// TIA Portal V21 export
// export: Created 2026-11-21T23:19:43.1672142Z, ExportSetting WithDefaults, DisplayName Totally Integrated Automation Portal, DisplayVersion V21 Update 3, DisplayName STEP 7 Professional, DisplayVersion V21 Update 3, DisplayName STEP 7 Safety, DisplayVersion V21, DisplayName Tech WebApplication, DisplayVersion V21, DisplayName WinCC Basic/Comfort/Advanced, DisplayVersion V21 Update 3, DisplayName WinCC Unified, DisplayVersion V21 Update 3
TagTable "Default tag table"
  Hmi_Bool : Bool  (1 s)
  Hmi_Int : Int  (1 s)
  Hmi_Real : Real  (1 s)
  Hmi_String : WString  (1 s)
  Ext_Bool : Bool  (PLC tag Plc_Bool, HMI_Connection_4, 1 s)
  Ext_Int : Int  (PLC tag Plc_Int, HMI_Connection_4, 1 s)
  Ext_Real : Real  (PLC tag Plc_Real, HMI_Connection_4, 1 s)
  Ext_Byte : Byte  (PLC tag Plc_Byte, HMI_Connection_4, 1 s)
